Yaskawa INFORM job: FEATURE.JBI

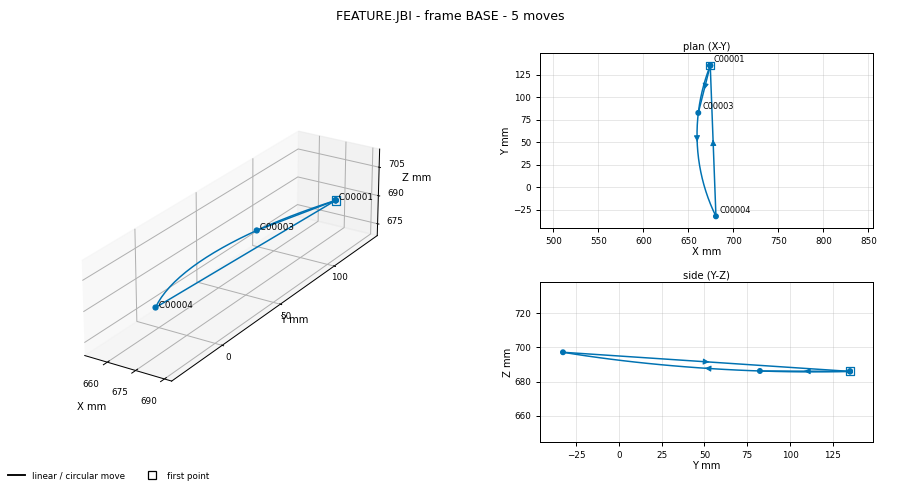
[picture p0: tool path of FEATURE.JBI in frame BASE, 5 of 8 moves have a stored position in this frame; points joined in program order, loops and branches not executed]
/JOB
//NAME FEATURE
//POS
///NPOS 8,0,0,0,0,0
///TOOL 1
///POSTYPE PULSE
///PULSE
C00000=10,20,-10,30,-45,60
///TOOL 1
///POSTYPE BASE
///RECTAN
///RCONF 0,0,0,0,0,0,0,0
C00001=674.300,134.999,685.980,-66.22,8.38,-107.67
C00002=674.300,134.999,685.980,-66.22,8.38,-107.67
C00003=661.027,82.386,686.221,-67.04,7.80,-111.79
C00004=680.634,-32.579,697.148,-65.39,8.96,-121.55
C00005=674.300,134.999,685.980,-66.22,8.38,-107.67
C00006=661.027,82.386,686.221,-67.04,7.80,-111.79
///POSTYPE PULSE
///PULSE
C00007=10,20,-10,30,-45,60
//INST
///DATE 2026/10/26 01:18
///COMM Generated using RoboDK
///ATTR SC,RW,RJ
///GROUP1 RB1
NOP
'Program generated by Vertical
'Bot Studio for Motoman GP8 on
' 25/10/2026 12:00:00
'Using nominal kinematics.
'Using Frame 2 (targets wrt ba
'se):
'100.0,-50.0,20.0,0.0,0.0,30.0
'Tool 1 (Tool 1) should be clo
'se to:
'10.0,0.0,120.0,0.0,15.0,0.0
MOVJ C00000 VJ=90.00
MOVL C00001 V=300.0
MOVC C00002 V=300.0 PL=5
MOVC C00003 V=300.0 PL=5
MOVC C00004 V=300.0 PL=5
MOVL C00005 V=50.0 ACC=100 DEC=100
MOVL C00006 V=300.0 ACC=100 DEC=100
DOUT OT#(3) ON
DOUT DO_GRIP OFF
WAIT IN#(5)=ON
WAIT DI_PART=ON T=2.00
TIMER T=0.50
'a comment line
MSG "Hello operator"
CALL JOB:MYFUNC
CALL JOB:SETRPM(
RAW_CODE_LINE
CALL JOB:SUBPICK
'Tool 1 (Tool 1) should be clo
'se to:
'10.0,0.0,120.0,0.0,15.0,0.0
'Attach to Tool 1
MOVJ C00007 VJ=45.00 ACC=100 DEC=100
PAUSE
END
